{region 'Documentation'}
(*!
<summary>Checks real Preparation-to-test handover; loss of Ready/Completed does not restart or block the active Test Case.</summary>
*)
{endregion}
FUNCTION_BLOCK Test_PreparationCompletionTracksTarget EXTENDS TestCaseBase
VAR
    FSubject : Prepare_ValueAtTarget;
    FResource : PreparationResource;
    FView : I_Preparation;
    FResourceAvailable : BOOL := TRUE;
    FObserved : ST_PreparationStatus;
    FExpected : ST_PreparationStatus;
    FObservedEnabled : BOOL;
    FExpectedEnabled : BOOL;
    FCheckPerformed : BOOL;
    FObservedCommandWrites : UDINT;
    FExpectedCommandWrites : UDINT;
    FObservedActualValue : DINT;
    FExpectedActualValue : DINT;
    FObservedRequestedValue : DINT;
    FExpectedRequestedValue : DINT;
    FCheckDiagnosticState : AssertEqual_Int;
    FCheckExecutionStatus : AssertEqual_Int;
    FCheckReady : AssertEqual_Bool;
    FCheckRunning : AssertEqual_Bool;
    FCheckCompleted : AssertEqual_Bool;
    FCheckError : AssertEqual_Bool;
    FCheckEnabled : AssertEqual_Bool;
    FCheckCommandWrites : AssertEqual_UDInt;
    FCheckActualValue : AssertEqual_DInt;
    FCheckRequestedValue : AssertEqual_DInt;
    FCheckTestingActive : AssertEqual_Bool;
END_VAR
VAR CONSTANT
    PreparationHandedOver : E_State := E_State.Running;
    TargetAndReadinessLost : E_State := E_State.Running + 1;
    TestingContinues : E_State := E_State.Running + 2;
END_VAR

SUPER^();

{region 'Documentation'}
(*!
<summary>Contributes all owned Assertion results without executing the subjects.</summary>
*)
{endregion}
METHOD PROTECTED AggregateResults
VAR_INPUT
    Aggregator : I_ResultAggregator; //! Borrowed result sink owned by the outer Test Case; add this test's checking Assertions without resetting or retaining the sink.
END_VAR
Aggregator.AddProvider(Provider := FCheckDiagnosticState);
Aggregator.AddProvider(Provider := FCheckExecutionStatus);
Aggregator.AddProvider(Provider := FCheckReady);
Aggregator.AddProvider(Provider := FCheckRunning);
Aggregator.AddProvider(Provider := FCheckCompleted);
Aggregator.AddProvider(Provider := FCheckError);
Aggregator.AddProvider(Provider := FCheckEnabled);
Aggregator.AddProvider(Provider := FCheckCommandWrites);
Aggregator.AddProvider(Provider := FCheckActualValue);
Aggregator.AddProvider(Provider := FCheckRequestedValue);
Aggregator.AddProvider(Provider := FCheckTestingActive);
END_METHOD

{region 'Documentation'}
(*!
<summary>Requires valid base configuration and every owned Assertion.</summary>
*)
{endregion}
METHOD PROTECTED CheckInitialization : BOOL //! TRUE when the inherited initialization check and this concrete fixture check both accept the setup.
CheckInitialization := FALSE;
IF NOT SUPER^.CheckInitialization() THEN
    RETURN;
END_IF;
IF NOT FCheckDiagnosticState.IsInitialized
    OR NOT FCheckExecutionStatus.IsInitialized
    OR NOT FCheckReady.IsInitialized
    OR NOT FCheckRunning.IsInitialized
    OR NOT FCheckCompleted.IsInitialized
    OR NOT FCheckError.IsInitialized
    OR NOT FCheckEnabled.IsInitialized
    OR NOT FCheckCommandWrites.IsInitialized
    OR NOT FCheckActualValue.IsInitialized
    OR NOT FCheckRequestedValue.IsInitialized
    OR NOT FCheckTestingActive.IsInitialized THEN
    RETURN;
END_IF;

CheckInitialization := TRUE;
END_METHOD

{region 'Documentation'}
(*!
<summary>Configures this scenario, its local subjects and named Assertions.</summary>
*)
{endregion}
METHOD PROTECTED Configure
FPreparationStateCount := 1;
FTestStateCount := 3;
FCheckPerformed := FALSE;
FResource.Initialize(InitialValue := 2);
FSubject.Initialize(Resource := FResource);
FView := FSubject;
FResourceAvailable := TRUE;

FCheckDiagnosticState.Initialize(Parent := THIS^,
    AssertionName := 'DiagnosticState');
FCheckExecutionStatus.Initialize(Parent := THIS^,
    AssertionName := 'ExecutionStatus');
FCheckReady.Initialize(Parent := THIS^,
    AssertionName := 'Ready');
FCheckRunning.Initialize(Parent := THIS^,
    AssertionName := 'Running');
FCheckCompleted.Initialize(Parent := THIS^,
    AssertionName := 'Completed');
FCheckError.Initialize(Parent := THIS^,
    AssertionName := 'Error');
FCheckEnabled.Initialize(Parent := THIS^,
    AssertionName := 'Enabled');
FCheckCommandWrites.Initialize(Parent := THIS^,
    AssertionName := 'CommandWrites');
FCheckActualValue.Initialize(Parent := THIS^,
    AssertionName := 'ActualValue');
FCheckRequestedValue.Initialize(Parent := THIS^,
    AssertionName := 'RequestedValue');
FCheckTestingActive.Initialize(Parent := THIS^,
    AssertionName := 'TestingActive');
END_METHOD

{region 'Documentation'}
(*!
<summary>Ends scenario processing without issuing further resource commands.</summary>
*)
{endregion}
METHOD PROTECTED ProcessAbort
VAR_INPUT
    Enable : BOOL; //! Phase permission supplied by the owning Test Case; FALSE does not authorize progression, while observation may continue.
END_VAR
IF Enable THEN
    CompleteAbort();
END_IF;
END_METHOD

{region 'Documentation'}
(*!
<summary>Compares independent expected values with the captured observations; called when disabled as well.</summary>
*)
{endregion}
METHOD PROTECTED ProcessAssertions
VAR_INPUT
    Enable : BOOL; //! Phase permission supplied by the owning Test Case; FALSE does not authorize progression, while observation may continue.
END_VAR
FCheckDiagnosticState(Enable := Enable,
    State := State,
    IN := TO_INT(FObserved.State),
    Expected := TO_INT(FExpected.State));

FCheckExecutionStatus(Enable := Enable,
    State := State,
    IN := TO_INT(FObserved.ExecutionStatus),
    Expected := TO_INT(FExpected.ExecutionStatus));

FCheckReady(Enable := Enable,
    State := State,
    IN := FObserved.Ready,
    Expected := FExpected.Ready);

FCheckRunning(Enable := Enable,
    State := State,
    IN := FObserved.Running,
    Expected := FExpected.Running);

FCheckCompleted(Enable := Enable,
    State := State,
    IN := FObserved.Completed,
    Expected := FExpected.Completed);

FCheckError(Enable := Enable,
    State := State,
    IN := FObserved.Error,
    Expected := FExpected.Error);

FCheckEnabled(Enable := Enable,
    State := State,
    IN := FObservedEnabled,
    Expected := FExpectedEnabled);

FCheckCommandWrites(Enable := Enable,
    State := State,
    IN := FObservedCommandWrites,
    Expected := FExpectedCommandWrites);

FCheckActualValue(Enable := Enable,
    State := State,
    IN := FObservedActualValue,
    Expected := FExpectedActualValue);

FCheckRequestedValue(Enable := Enable,
    State := State,
    IN := FObservedRequestedValue,
    Expected := FExpectedRequestedValue);

FCheckTestingActive(Enable := Enable,
    State := State,
    IN := IsTestingActive,
    Expected := TRUE);

IF Enable
    AND FCheckDiagnosticState.EvaluationActive
    AND FCheckExecutionStatus.EvaluationActive
    AND FCheckReady.EvaluationActive
    AND FCheckRunning.EvaluationActive
    AND FCheckCompleted.EvaluationActive
    AND FCheckError.EvaluationActive
    AND FCheckEnabled.EvaluationActive
    AND FCheckCommandWrites.EvaluationActive
    AND FCheckActualValue.EvaluationActive
    AND FCheckRequestedValue.EvaluationActive
    AND FCheckTestingActive.EvaluationActive THEN
    FCheckPerformed := TRUE;
END_IF;
END_METHOD

{region 'Documentation'}
(*!
<summary>Runs the real Preparation phase and projects its observations to the owner.</summary>
*)
{endregion}
METHOD PROTECTED ProcessPreparations
VAR_INPUT
    Enable : BOOL; //! Phase permission supplied by the owning Test Case; FALSE does not authorize progression, while observation may continue.
END_VAR
FResource(Available := FResourceAvailable,
    Fault := FALSE,
    Advance := TRUE);
FSubject(Enable := Enable,
    TargetValue := 0);
FObserved := FView.Status;
UpdatePreparationStatus(Ready := FObserved.Ready,
    Running := FObserved.Running,
    Completed := FObserved.Completed,
    HasError := FObserved.Error,
    State := FObserved.State);
END_METHOD

{region 'Documentation'}
(*!
<summary>Restores repeatable fixture state and resets Assertions before returning to Idle.</summary>
*)
{endregion}
METHOD PROTECTED ProcessReset
FCheckPerformed := FALSE;
FResource.Initialize(InitialValue := 2);
FSubject.Initialize(Resource := FResource);
FView := FSubject;
FResourceAvailable := TRUE;
FCheckDiagnosticState.Reset();
FCheckExecutionStatus.Reset();
FCheckReady.Reset();
FCheckRunning.Reset();
FCheckCompleted.Reset();
FCheckError.Reset();
FCheckEnabled.Reset();
FCheckCommandWrites.Reset();
FCheckActualValue.Reset();
FCheckRequestedValue.Reset();
FCheckTestingActive.Reset();
CompleteReset();
END_METHOD

{region 'Documentation'}
(*!
<summary>Exercises one named scenario step per call; advances only after actual Assertion evaluation.</summary>
*)
{endregion}
METHOD PROTECTED ProcessTests
VAR_INPUT
    Enable : BOOL; //! Phase permission supplied by the owning Test Case; FALSE does not authorize progression, while observation may continue.
END_VAR
IF NOT Enable THEN
    RETURN;
END_IF;

IF FCheckPerformed THEN
    FCheckPerformed := FALSE;
    IF State = TestingContinues THEN
        CompleteTests();
        RETURN;
    END_IF;
    NextTestState();
    IF NOT IsTestingActive THEN
        RETURN;
    END_IF;
END_IF;

CASE State OF
    PreparationHandedOver:
        FResource.RequestValue(Value := 2);
        FResourceAvailable := FALSE;
        FExpected.State := E_State.Completed;
        FExpected.ExecutionStatus := E_ExecutionStatus.Completed;
        FExpected.Ready := TRUE;
        FExpected.Running := FALSE;
        FExpected.Completed := TRUE;
        FExpected.Error := FALSE;
        FExpectedEnabled := FALSE;
        FExpectedCommandWrites := 2;
        FExpectedActualValue := 0;
        FExpectedRequestedValue := 2;

    TargetAndReadinessLost:
        FExpected.State := E_State.Idle;
        FExpected.ExecutionStatus := E_ExecutionStatus.NotReady;
        FExpected.Ready := FALSE;
        FExpected.Running := FALSE;
        FExpected.Completed := FALSE;
        FExpected.Error := FALSE;
        FExpectedEnabled := FALSE;
        FExpectedCommandWrites := 2;
        FExpectedActualValue := 0;
        FExpectedRequestedValue := 2;

    TestingContinues:
        FExpected.State := E_State.Idle;
        FExpected.ExecutionStatus := E_ExecutionStatus.NotReady;
        FExpected.Ready := FALSE;
        FExpected.Running := FALSE;
        FExpected.Completed := FALSE;
        FExpected.Error := FALSE;
        FExpectedEnabled := FALSE;
        FExpectedCommandWrites := 2;
        FExpectedActualValue := 0;
        FExpectedRequestedValue := 2;

ELSE
    Error(Message := 'Unexpected Preparation test state.');
    RETURN;
END_CASE;

FObserved := FView.Status;
FObservedEnabled := FSubject.Enabled;

FObservedCommandWrites := FResource.CommandWriteCount;
FObservedActualValue := FResource.ActualValue;
FObservedRequestedValue := FResource.RequestedValue;
END_METHOD

END_FUNCTION_BLOCK

(* stored: Version 1.1.0.1
   POU Test_PreparationCompletionTracksTarget: Id {6b1f7926-3bfe-4c7e-bc3e-aae8b157270c}, SpecialFunc None
   Folder Internal: Id {77bf36f8-8426-427e-9fea-9d664f340270}
   Method AggregateResults: Id {38033f6b-1a27-4b67-aed4-a72e1dcdc379}
   Method CheckInitialization: Id {392f05f5-19a8-4080-ae00-905f7ea81998}
   Method Configure: Id {ae0235f2-f6b9-4463-9cbe-c87321119595}
   Method ProcessAbort: Id {fcfc41d1-6b58-479f-a0ca-97d3ef37fd52}
   Method ProcessAssertions: Id {d35485c2-10cb-4589-b112-4b48963ad4ca}
   Method ProcessPreparations: Id {04d5786b-21d3-41f2-94bf-cb4cb6670d86}
   Method ProcessReset: Id {c93c2117-91db-4c4e-ad02-e053d49be423}
   Method ProcessTests: Id {9d5dcddb-844d-450d-af85-3300a6466918} *)
